// TIA Portal V20 export
Screen "Pop-up_Opmodes6_Popup"  645x267
  ScreenItem "Background" at 0,0 size 645x267  Type=HmiRectangle
  ScreenItem "Descr_HmiPanel" at 1,208 size 56x40  Type=HmiTextBox
  ScreenItem "Linie1_LightGrey" at 10,207 size 520x0  Type=HmiLine
  ScreenItem "Linie1_DarkGrey" at 10,207 size 520x0  Type=HmiLine
  ScreenItem "Linie1_LightGrey_1" at 10,249 size 520x0  Type=HmiLine
  ScreenItem "Linie1_DarkGrey_1" at 10,248 size 520x0  Type=HmiLine
  ScreenItem "Overview_OPMode" at 1,1 size 643x25  Type=HmiTextBox
  ScreenItem "Descr_OPMode" at 1,26 size 550x40  Type=HmiTextBox
  ScreenItem "OPMode1_small" at 13,104 size 90x60  Type=HmiButton
  ScreenItem "OPMode2_small" at 120,104 size 90x60  Type=HmiButton
  ScreenItem "OPMode3_small" at 226,104 size 90x60  Type=HmiButton
  ScreenItem "OPMode5_small" at 439,104 size 90x60  Type=HmiButton
  ScreenItem "OPMode4_small" at 333,104 size 90x60  Type=HmiButton
  ScreenItem "OPMode6_small" at 545,104 size 90x60  Type=HmiButton
  ScreenItem "OPMode1_wide" at 8,104 size 100x60  Type=HmiButton
  ScreenItem "OPMode2_wide" at 115,104 size 100x60  Type=HmiButton
  ScreenItem "OPMode3_wide" at 221,104 size 100x60  Type=HmiButton
  ScreenItem "OPMode4_wide" at 327,104 size 100x60  Type=HmiButton
  ScreenItem "OPMode5_wide" at 434,104 size 100x60  Type=HmiButton
  ScreenItem "OPMode6_wide" at 540,104 size 100x60  Type=HmiButton
  ScreenItem "Overview_HMI-OP" at 554,207 size 90x60  Type=HmiButton
  ScreenItem "Cancel Mode" at 554,1 size 90x60  Type=HmiButton
  ScreenItem "OPMode1_Foreground_Blocked" at 7,104 size 100x60  Type=HmiGraphicView
  ScreenItem "OPMode2_Foreground_Blocked" at 112,104 size 100x60  Type=HmiGraphicView
  ScreenItem "OPMode3_Foreground_Blocked" at 219,104 size 100x60  Type=HmiGraphicView
  ScreenItem "OPMode4_Foreground_Blocked" at 327,104 size 100x60  Type=HmiGraphicView
  ScreenItem "OPMode5_Foreground_Blocked" at 434,104 size 100x60  Type=HmiGraphicView
  ScreenItem "OPMode6_Foreground_Blocked" at 540,104 size 100x60  Type=HmiGraphicView
  ScreenItem "OPMode1_Blocked" at 93,106 size 14x14  Type=HmiGraphicView
  ScreenItem "OPMode2_Blocked" at 200,106 size 14x14  Type=HmiGraphicView
  ScreenItem "OPMode3_Blocked" at 305,106 size 14x14  Type=HmiGraphicView
  ScreenItem "OPMode4_Blocked" at 411,106 size 14x14  Type=HmiGraphicView
  ScreenItem "OPMode5_Blocked" at 518,106 size 14x14  Type=HmiGraphicView
  ScreenItem "OPMode6_Blocked" at 625,106 size 14x14  Type=HmiGraphicView
